--- program BumperF_C (robot ABB IRB 1300-10/1.15) ---
  Smooth(1)
  Set speed (1000.0 mm/s)
  Set Ref.: BumperF
  Set Tool: Generic Paint Sprayer
  Show Generic Paint Sprayer
  MoveJ 1 to (1571.24, -957.53, 569.46) mm, rotated rx 115.95 ry -6.64 rz -166.63 deg; joints [132.246, 136.209, -181.396, 156.344, 105.383, -115.772, 4593.947, 921.715, 1041.563]
  MoveL 2 to (1571.24, -957.53, 569.46) mm, rotated rx 115.95 ry -6.64 rz -166.63 deg; joints [132.246, 136.209, -181.396, 156.344, 105.383, -115.772, 4593.947, 921.715, 1041.563]
  MoveL 3 to (1545.53, -871.22, 525.99) mm, rotated rx 115.95 ry -6.64 rz -166.63 deg; joints [132.246, 136.209, -181.396, 156.344, 105.383, -115.772, 4568.236, 1008.026, 1085.031]
  MoveL 4 to (1545.53, -871.22, 525.99) mm, rotated rx 115.95 ry -6.64 rz -166.63 deg; joints [132.246, 136.209, -181.396, 156.344, 105.383, -115.772, 4568.236, 1008.026, 1085.031]
  Set speed (200.0 mm/s)
  MoveL 5 to (1567.25, -870.44, 513.69) mm, rotated rx 114.53 ry -6.57 rz -165.92 deg; joints [131.765, 135.013, -181.396, 155.74, 105.383, -114.904, 4591.602, 1008.066, 1094.602]
  MoveL 6 to (1592.89, -869.13, 497.74) mm, rotated rx 110.93 ry -5.65 rz -165.57 deg; joints [130.698, 131.085, -181.396, 155.714, 105.383, -112.016, 4607.617, 1008.267, 1096.076]
  MoveL 7 to (1616.69, -868.87, 477.59) mm, rotated rx 107.37 ry -5.12 rz -164.07 deg; joints [129.332, 127.093, -181.396, 154.983, 104.902, -109.292, 4628.08, 1008.268, 1100]
  MoveL 8 to (1638.67, -867.82, 457.97) mm, rotated rx 105.23 ry -4.69 rz -163.28 deg; joints [128.5, 123.788, -181.396, 154.835, 103.912, -107.249, 4645.228, 1008.269, 1099.981]
  MoveL 9 to (1659.86, -866.51, 437.3) mm, rotated rx 104.04 ry -4.24 rz -163.53 deg; joints [128.5, 121.033, -181.396, 155.103, 102.7, -105.772, 4660.763, 1003.997, 1100]
  MoveL 10 to (1680.53, -864.68, 416.9) mm, rotated rx 102.62 ry -4.06 rz -162.44 deg; joints [127.494, 118.2, -181.396, 154.969, 101.395, -104.09, 4676.396, 1006.029, 1100]
  MoveL 11 to (1700.41, -862.07, 396.49) mm, rotated rx 100.96 ry -3.66 rz -161.77 deg; joints [126.76, 115.027, -181.132, 154.969, 100.379, -102.383, 4689.707, 1006.022, 1100]
  MoveL 12 to (1721.6, -858.14, 377.92) mm, rotated rx 98.48 ry -2.82 rz -161.72 deg; joints [126.547, 111.062, -179.997, 154.969, 100.379, -100.648, 4704.908, 1003.768, 1100]
  MoveL 13 to (1729.97, -859.97, 342.08) mm, rotated rx 96.18 ry -2.12 rz -161.17 deg; joints [125.885, 105.454, -176.974, 154.97, 100.379, -99.014, 4709.436, 1003.105, 1100]
  MoveL 14 to (1729.45, -862.07, 324.55) mm, rotated rx 95.53 ry -1.83 rz -161.71 deg; joints [126.39, 103.099, -175.393, 154.981, 100.379, -98.605, 4709.436, 996.85, 1100]
  MoveL 15 to (1734.68, -862.07, 305.71) mm, rotated rx 94.94 ry -1.6 rz -162.14 deg; joints [126.39, 100.689, -173.732, 155.4, 100.379, -98.09, 4710.155, 996.383, 1100]
  MoveL 16 to (1743.31, -860.76, 287.4) mm, rotated rx 94.35 ry -1.49 rz -161.17 deg; joints [125.481, 98.526, -173.288, 155.4, 99.369, -97.19, 4712.272, 996.382, 1100]
  MoveL 17 to (1754.56, -857.88, 271.44) mm, rotated rx 93.88 ry -1.28 rz -161.73 deg; joints [125.481, 96.542, -172.176, 155.976, 99.142, -96.642, 4715.904, 996.382, 1100]
  MoveL 18 to (1759.01, -858.14, 245.02) mm, rotated rx 92.82 ry -0.95 rz -161.34 deg; joints [125.066, 92.989, -169.805, 155.975, 99.142, -95.921, 4715.904, 993.682, 1100]
  MoveL 19 to (1756.13, -859.71, 226.97) mm, rotated rx 92.24 ry -0.73 rz -162.03 deg; joints [125.745, 90.661, -168.159, 155.976, 99.142, -95.55, 4711.513, 983.719, 1100]
  MoveL 20 to (1756.92, -860.24, 208.39) mm, rotated rx 91.53 ry -0.48 rz -162.48 deg; joints [126.192, 88.179, -166.477, 155.976, 99.142, -95.085, 4709.215, 974.937, 1100]
  MoveL 21 to (1757.7, -860.24, 190.6) mm, rotated rx 91.06 ry -0.32 rz -163.42 deg; joints [127.122, 85.976, -164.811, 155.976, 99.142, -94.779, 4708.177, 964.459, 1100]
  MoveL 22 to (1758.49, -860.24, 174.38) mm, rotated rx 90.59 ry -0.18 rz -163.41 deg; joints [127.122, 83.931, -163.287, 155.969, 99.142, -94.457, 4705.559, 959.867, 1100]
  MoveL 23 to (1758.75, -860.24, 159.73) mm, rotated rx 90.12 ry -0.03 rz -163.88 deg; joints [127.59, 82.032, -161.91, 155.969, 99.142, -94.134, 4702.574, 951.798, 1100]
  MoveL 24 to (1759.27, -859.97, 146.91) mm, rotated rx 90 ry 0 rz -165.53 deg; joints [129.218, 80.632, -160.641, 155.988, 99.142, -94.048, 4702.574, 938.888, 1100]
  MoveL 25 to (1760.58, -859.71, 136.45) mm, rotated rx 90.12 ry -0.04 rz -162.94 deg; joints [127.222, 79.74, -160.641, 155.454, 98.168, -93.794, 4702.575, 945.045, 1099.999]
  MoveL 26 to (1763.2, -858.93, 129.12) mm, rotated rx 90.71 ry -0.2 rz -164.47 deg; joints [128.117, 79.543, -159.846, 156.101, 98.168, -94.096, 4702.574, 944.116, 1100]
  Set speed (1000.0 mm/s)
  MoveL 27 to (1763.2, -858.93, 129.12) mm, rotated rx 90.71 ry -0.2 rz -164.47 deg; joints [128.117, 79.543, -159.846, 156.101, 98.168, -94.096, 4702.574, 944.116, 1100]
  MoveL 28 to (1789.97, -955.27, 130.36) mm, rotated rx 90.71 ry -0.2 rz -164.47 deg; joints [128.117, 79.543, -159.846, 156.101, 98.168, -94.096, 4729.346, 847.775, 1098.767]
  Set speed (1000.0 mm/s)
  MoveL 29 to (1779.18, -953.4, 138.35) mm, rotated rx 98.16 ry 0.3 rz 177.94 deg; joints [138.476, 85.541, -159.846, 163.825, 98.168, -98.714, 4697.875, 847.774, 1094.184]
  MoveL 30 to (1782.82, -854.48, 124.15) mm, rotated rx 98.16 ry 0.3 rz 177.94 deg; joints [138.575, 84.798, -159.846, 163.754, 97.448, -98.53, 4697.874, 941.635, 1100]
  MoveL 31 to (1782.82, -854.48, 124.15) mm, rotated rx 98.16 ry 0.3 rz 177.94 deg; joints [138.575, 84.798, -159.846, 163.754, 97.448, -98.53, 4697.874, 941.635, 1100]
  Set speed (200.0 mm/s)
  MoveL 32 to (1786.22, -852.91, 135.66) mm, rotated rx 96.28 ry 0.04 rz 179.68 deg; joints [137.268, 84.574, -160.749, 163.124, 97.823, -97.175, 4697.874, 941.635, 1100]
  MoveL 33 to (1790.67, -851.08, 147.7) mm, rotated rx 98.11 ry -0.22 rz -178.44 deg; joints [135.583, 84.574, -160.749, 163.124, 96.101, -97.893, 4702.805, 954.913, 1071.274]
  MoveL 34 to (1796.68, -848.72, 159.47) mm, rotated rx 98.74 ry -0.53 rz -176.58 deg; joints [133.77, 84.574, -160.749, 163.124, 95.404, -97.953, 4707.715, 968.876, 1052.965]
  MoveL 35 to (1802.7, -846.37, 171.77) mm, rotated rx 98.62 ry -0.68 rz -175.51 deg; joints [133.516, 84.592, -160.749, 162.287, 95.39, -97.953, 4720.878, 970.014, 1041.305]
  MoveL 36 to (1809.24, -843.75, 184.32) mm, rotated rx 99.8 ry -0.99 rz -174.27 deg; joints [132.393, 84.592, -160.749, 162.287, 94.205, -98.297, 4727.536, 980.866, 1017.452]
  MoveL 37 to (1816.57, -840.61, 197.4) mm, rotated rx 100.78 ry -1.11 rz -174.17 deg; joints [132.393, 84.592, -160.749, 162.298, 93.3, -98.698, 4735.96, 985.217, 995.643]
  MoveL 38 to (1824.41, -837.21, 211.01) mm, rotated rx 101.64 ry -1.18 rz -174.28 deg; joints [132.393, 84.592, -160.749, 162.521, 92.536, -99.039, 4742.893, 990.437, 974.508]
  MoveL 39 to (1824.41, -837.21, 211.01) mm, rotated rx 93.53 ry -1.19 rz -161.37 deg; joints [123.735, 79.476, -160.749, 157.598, 94.418, -94.055, 4742.893, 990.436, 988.777]
  MoveL 40 to (1820.23, -837.21, 231.94) mm, rotated rx 93.35 ry -1.2 rz -160.31 deg; joints [123.243, 79.476, -160.872, 157.02, 94.418, -93.99, 4742.894, 992.111, 969.266]
  MoveL 41 to (1820.23, -837.21, 231.94) mm, rotated rx 101.71 ry -1.43 rz -173.11 deg; joints [131.794, 84.617, -160.872, 161.941, 92.215, -98.959, 4742.894, 992.113, 952.179]
  MoveL 42 to (1829.38, -833.03, 246.59) mm, rotated rx 102.88 ry -1.89 rz -171.78 deg; joints [130.559, 84.617, -160.872, 161.941, 90.966, -99.177, 4752.022, 1006.027, 925.876]
  MoveL 43 to (1839.06, -828.32, 260.98) mm, rotated rx 103.06 ry -1.91 rz -171.82 deg; joints [130.559, 84.617, -160.872, 162.004, 90.806, -99.242, 4761.37, 1011.202, 909.915]
  MoveL 44 to (1849.01, -823.35, 275.1) mm, rotated rx 104.57 ry -2.33 rz -171.12 deg; joints [130.013, 84.617, -160.872, 162.004, 89.294, -99.68, 4772.697, 1022.45, 881.62]
  MoveL 45 to (1863.66, -815.76, 294.46) mm, rotated rx 107.07 ry -3 rz -170.32 deg; joints [129.479, 84.698, -160.872, 162.004, 86.864, -100.462, 4790.854, 1039.487, 839.866]
  MoveL 46 to (1882.49, -804.77, 317.22) mm, rotated rx 109.65 ry -4.19 rz -168.43 deg; joints [127.743, 84.698, -160.872, 162.004, 84.028, -100.823, 4811.061, 1068.912, 791.558]
  MoveL 47 to (1895.83, -796.14, 330.83) mm, rotated rx 113.34 ry -6.41 rz -165.49 deg; joints [124.807, 84.698, -160.872, 162.004, 79.723, -100.879, 4824.82, 1109.926, 740.477]
  MoveL 48 to (1904.47, -789.86, 337.89) mm, rotated rx 116.65 ry -8.76 rz -163.11 deg; joints [122.23, 85.616, -160.872, 162.003, 76.566, -100.879, 4837.457, 1154.33, 710.031]
  MoveL 49 to (1913.1, -783.32, 343.38) mm, rotated rx 120.5 ry -11.96 rz -160.62 deg; joints [119.262, 88.097, -160.872, 162.003, 74.023, -100.879, 4855.125, 1218.718, 694.119]
  MoveL 50 to (1922, -776, 347.57) mm, rotated rx 123.01 ry -13.87 rz -159.75 deg; joints [118.011, 89.326, -160.872, 162.003, 72.107, -100.879, 4869.128, 1258.002, 680.927]
  MoveL 51 to (1931.15, -768.41, 350.45) mm, rotated rx 127.02 ry -16.88 rz -158.94 deg; joints [116.434, 91.393, -160.872, 162.003, 69.207, -100.88, 4887.234, 1316.61, 667.809]
  MoveL 52 to (1940.57, -759.78, 352.02) mm, rotated rx 133.81 ry -20.92 rz -159.59 deg; joints [115.619, 92.398, -160.872, 162.003, 62.545, -100.88, 4909.28, 1386.174, 628.482]
  MoveL 53 to (1949.99, -750.62, 352.54) mm, rotated rx 133.85 ry -22.45 rz -158.32 deg; joints [113.518, 92.645, -160.872, 161.597, 62.116, -99.201, 4909.281, 1414.858, 628.482]
  MoveL 54 to (1959.93, -740.68, 352.54) mm, rotated rx 138.13 ry -26.48 rz -158.22 deg; joints [110.548, 94.884, -160.872, 161.597, 59.126, -97.312, 4911.466, 1494.181, 628.482]
  MoveL 55 to (1970.13, -729.69, 351.76) mm, rotated rx 138.94 ry -28.75 rz -157.27 deg; joints [108.289, 95.245, -160.871, 160.752, 58.015, -95.019, 4911.466, 1532.276, 628.482]
  MoveL 56 to (1980.07, -718.44, 350.97) mm, rotated rx 138.97 ry -29.76 rz -156.64 deg; joints [106.869, 95.245, -160.871, 160.411, 57.708, -93.633, 4911.467, 1554.428, 628.83]
  MoveL 57 to (1989.75, -706.93, 349.92) mm, rotated rx 136.16 ry -29.58 rz -154.64 deg; joints [105.639, 94.385, -160.871, 159.72, 59.288, -92.34, 4911.466, 1550.094, 633.425]
  MoveL 58 to (1998.91, -695.68, 349.4) mm, rotated rx 133.19 ry -28.72 rz -152.89 deg; joints [104.809, 93.375, -160.871, 159.442, 61.115, -91.65, 4911.467, 1539.501, 637.871]
  MoveL 59 to (2007.02, -685.48, 349.66) mm, rotated rx 130.86 ry -27.24 rz -152.11 deg; joints [104.689, 92.218, -160.872, 159.777, 62.539, -91.731, 4911.472, 1524.592, 637.872]
  MoveL 60 to (2014.35, -675.8, 350.97) mm, rotated rx 122.46 ry -23.36 rz -148.07 deg; joints [103.96, 90.632, -160.872, 159.151, 69.542, -91.731, 4911.472, 1473.431, 675.241]
  MoveL 61 to (2038.15, -649.11, 345.74) mm, rotated rx 114.17 ry -24.24 rz -137.55 deg; joints [97.018, 85.715, -160.872, 155.117, 71.4, -85.824, 4911.471, 1473.426, 679.245]
  MoveL 62 to (2051.49, -633.42, 343.12) mm, rotated rx 112.8 ry -23.19 rz -136.86 deg; joints [96.789, 84.623, -160.872, 155.117, 71.99, -85.767, 4922.042, 1473.425, 681.907]
  MoveL 63 to (2063.79, -619.03, 341.03) mm, rotated rx 110.74 ry -21.37 rz -136.1 deg; joints [96.739, 82.665, -160.872, 155.117, 72.722, -85.767, 4931.522, 1459.566, 682.288]
  MoveL 64 to (2075.04, -605.69, 338.68) mm, rotated rx 110.8 ry -22.47 rz -134.83 deg; joints [94.985, 82.747, -160.872, 155.117, 72.306, -84.714, 4932.35, 1484.471, 682.288]
  MoveL 65 to (2085.24, -593.13, 336.58) mm, rotated rx 111.8 ry -23.63 rz -134.94 deg; joints [94.569, 83.495, -160.872, 155.119, 71.667, -84.319, 4940.301, 1511.538, 682.287]
  MoveL 66 to (2094.4, -581.62, 334.49) mm, rotated rx 111.31 ry -24.25 rz -133.53 deg; joints [92.994, 83.3, -160.872, 155.016, 71.667, -83.386, 4940.301, 1528.356, 684.409]
  MoveL 67 to (2102.51, -570.63, 332.4) mm, rotated rx 109.4 ry -23.08 rz -131.93 deg; joints [92.04, 82.56, -160.874, 155.016, 73.082, -83.386, 4943.467, 1528.189, 695.451]
  MoveL 68 to (2110.1, -560.43, 330.04) mm, rotated rx 108.78 ry -24.16 rz -129.72 deg; joints [90.063, 82.505, -160.874, 154.429, 73.082, -82.108, 4943.467, 1549.13, 699.124]
  MoveL 69 to (2116.64, -550.75, 327.16) mm, rotated rx 108.04 ry -24.56 rz -128.09 deg; joints [88.633, 82.011, -160.874, 154.121, 73.082, -81.209, 4943.468, 1560.135, 701.179]
  MoveL 70 to (2122.13, -542.64, 323.24) mm, rotated rx 107.35 ry -27.97 rz -123.66 deg; joints [85.357, 82.011, -160.874, 151.788, 72.164, -77.874, 4943.468, 1597.347, 702.069]
  MoveL 71 to (2126.32, -536.1, 317.48) mm, rotated rx 104.82 ry -29.37 rz -118.34 deg; joints [82.164, 80.426, -160.874, 149.535, 72.164, -74.977, 4943.468, 1609.549, 706.168]
  MoveL 72 to (2128.93, -531.65, 312.25) mm, rotated rx 101.45 ry -27.26 rz -113.85 deg; joints [79.937, 78.849, -160.874, 148.686, 74.318, -74.977, 4943.468, 1602.173, 725.352]
  MoveL 73 to (2128.93, -531.65, 312.25) mm, rotated rx 126.84 ry -33.58 rz -143.56 deg; joints [92.503, 91.12, -160.874, 157.962, 63.217, -81.642, 4943.468, 1719.806, 680.931]
  MoveL 74 to (2132.86, -524.59, 312.51) mm, rotated rx 131.8 ry -39.39 rz -144.63 deg; joints [90.442, 93.308, -160.873, 155.312, 59.914, -77.41, 4943.469, 1794.525, 680.931]
  MoveL 75 to (2138.61, -511.5, 310.94) mm, rotated rx 142.1 ry -48.23 rz -149.86 deg; joints [88.012, 93.628, -151.887, 151.963, 59.913, -73.067, 4943.469, 1959.558, 680.933]
  MoveL 76 to (2145.41, -491.62, 307.54) mm, rotated rx 148.42 ry -53.14 rz -153.81 deg; joints [86.275, 93.628, -151.373, 148.126, 56.76, -67.236, 4943.47, 2030.159, 680.933]
  MoveL 77 to (2152.48, -464.94, 303.62) mm, rotated rx 151.46 ry -56.88 rz -155.51 deg; joints [84.483, 93.628, -151.372, 144.702, 55.943, -62.304, 4943.47, 2082.544, 691.657]
  MoveL 78 to (2159.28, -432.5, 300.48) mm, rotated rx 157.96 ry -60.16 rz -160.65 deg; joints [83.237, 93.628, -150.316, 141.632, 54.856, -57.784, 4943.47, 2154.516, 700.89]
  MoveL 79 to (2166.08, -389.07, 298.39) mm, rotated rx 162.71 ry -60.68 rz -164.82 deg; joints [83.006, 93.628, -148.348, 141.49, 54.655, -57.243, 4943.475, 2227.842, 705.926]
  MoveL 80 to (2172.36, -330.47, 297.08) mm, rotated rx 166.98 ry -61.73 rz -168.49 deg; joints [82.432, 93.628, -147.038, 140.505, 54.605, -55.672, 4943.475, 2310.718, 713.199]
  MoveL 81 to (2178.12, -262.97, 296.29) mm, rotated rx 166.1 ry -61.33 rz -167.75 deg; joints [82.2, 93.628, -147.375, 141.056, 54.605, -55.884, 4943.475, 2371.713, 711.376]
  MoveL 82 to (2182.83, -193.12, 295.77) mm, rotated rx 169.21 ry -61.46 rz -170.5 deg; joints [82.021, 93.628, -146.721, 140.72, 54.052, -55.086, 4943.475, 2456.324, 712.371]
  MoveL 83 to (2185.96, -124.84, 295.51) mm, rotated rx 172.94 ry -62.25 rz -173.75 deg; joints [81.639, 93.628, -145.665, 139.712, 54.052, -53.733, 4943.475, 2544.405, 718.894]
  MoveL 84 to (2187.8, -61.27, 295.51) mm, rotated rx 174.69 ry -62.34 rz -175.3 deg; joints [81.557, 93.628, -144.992, 139.539, 54.052, -53.476, 4943.475, 2618.074, 721.416]
  MoveL 85 to (2189.1, -0.05, 295.51) mm, rotated rx -177.26 ry -62.45 rz 177.57 deg; joints [81.557, 93.628, -143.265, 137.966, 52.878, -51.455, 4943.475, 2717.714, 728.542]
  MoveL 86 to (2187.8, 61.17, 295.51) mm, rotated rx -173.75 ry -62.29 rz 174.47 deg; joints [81.71, 93.628, -142.223, 137.399, 52.478, -50.92, 4943.474, 2797.79, 733.234]
  MoveL 87 to (2185.96, 124.74, 295.51) mm, rotated rx -170.29 ry -62.04 rz 171.41 deg; joints [81.906, 93.628, -140.949, 136.945, 52.22, -50.617, 4943.472, 2881.625, 739.388]
  MoveL 88 to (2182.83, 193.28, 295.77) mm, rotated rx -166.22 ry -61.1 rz 167.88 deg; joints [82.416, 93.628, -139.453, 136.732, 51.343, -50.616, 4943.472, 2975.922, 744.195]
  MoveL 89 to (2178.12, 262.87, 296.29) mm, rotated rx -163.59 ry -60.95 rz 165.56 deg; joints [82.676, 93.628, -138.26, 136.285, 51.343, -50.526, 4943.472, 3062.322, 751.37]
  MoveL 90 to (2172.36, 330.37, 297.08) mm, rotated rx -163.15 ry -61.13 rz 165.14 deg; joints [82.913, 93.628, -138.152, 135.936, 51.343, -50.479, 4943.471, 3131.981, 752.579]
  MoveL 91 to (2166.08, 388.97, 298.39) mm, rotated rx -155.06 ry -58.82 rz 158.3 deg; joints [83.805, 93.628, -134.575, 135.497, 49.863, -50.479, 4943.471, 3246.959, 770.044]
  MoveL 92 to (2159.28, 432.4, 300.48) mm, rotated rx -150.95 ry -57.83 rz 154.82 deg; joints [84.274, 93.628, -132.455, 135.037, 49.517, -50.479, 4943.457, 3320.012, 783.091]
  MoveL 93 to (2152.48, 465.1, 303.62) mm, rotated rx -144.6 ry -53.45 rz 150.28 deg; joints [85.716, 93.628, -130.007, 135.037, 45.48, -50.342, 4943.456, 3409.512, 793.219]
  MoveL 94 to (2145.41, 491.52, 307.54) mm, rotated rx -142.77 ry -49.52 rz 149.98 deg; joints [86.332, 93.736, -130.007, 136.122, 41.249, -50.342, 4923.205, 3464.712, 785.161]
  MoveL 95 to (2138.61, 511.67, 310.94) mm, rotated rx -140.46 ry -46.77 rz 148.98 deg; joints [87.496, 93.756, -129.75, 136.122, 37.777, -50.276, 4923.205, 3511.087, 785.16]
  MoveL 96 to (2132.86, 524.49, 312.51) mm, rotated rx -133.08 ry -41.17 rz 144.86 deg; joints [88.774, 93.756, -125.065, 136.122, 33.797, -50.263, 4923.205, 3605.485, 833.592]
  MoveL 97 to (2128.93, 531.55, 312.25) mm, rotated rx -126.84 ry -33.58 rz 143.56 deg; joints [90.862, 93.756, -122.789, 136.122, 25.461, -49.709, 4923.205, 3689.917, 878.711]
  MoveL 98 to (2128.93, 531.55, 312.25) mm, rotated rx -100.25 ry -7.61 rz 109.92 deg; joints [121.937, 78.369, -126.316, 15.017, 36.087, 78.198, 5588.694, 3468.859, 878.521]
  MoveL 99 to (2126.32, 536, 317.48) mm, rotated rx -104.1 ry -29.19 rz 117.26 deg; joints [117.367, 96.341, -169.247, 16.72, 48.145, 64.164, 5423.205, 3346.609, 878.683]
  MoveL 100 to (2122.13, 542.54, 323.24) mm, rotated rx -105.97 ry -28.47 rz 120.97 deg; joints [117.367, 96.341, -169.247, 12.679, 46.638, 66.806, 5394.89, 3369.672, 861.092]
  MoveL 101 to (2116.64, 550.65, 327.16) mm, rotated rx -107.55 ry -25.57 rz 126.23 deg; joints [117.365, 96.872, -169.247, 5.15, 45.601, 72.802, 5349.984, 3412.333, 858.641]
  MoveL 102 to (2110.1, 560.33, 330.04) mm, rotated rx -108.36 ry -23.05 rz 130.28 deg; joints [117.365, 97.148, -169.622, -1.121, 45.94, 77.838, 5308.188, 3445.265, 858.641]
  MoveL 103 to (2102.51, 570.53, 332.4) mm, rotated rx -108.16 ry -21.99 rz 131.22 deg; joints [117.365, 97.148, -169.622, -2.931, 46.544, 79.449, 5290.898, 3463.725, 860.533]
  MoveL 104 to (2094.4, 581.52, 334.49) mm, rotated rx -112.03 ry -24.25 rz 134.57 deg; joints [117.365, 97.148, -169.622, -4.906, 42.427, 79.382, 5264.861, 3465.093, 824.183]
  MoveL 105 to (2085.24, 593.29, 336.58) mm, rotated rx -112.13 ry -23.27 rz 135.83 deg; joints [117.365, 97.206, -169.702, -7.138, 42.788, 81.232, 5243.276, 3484.334, 824.183]
  MoveL 106 to (2075.04, 605.59, 338.68) mm, rotated rx -109.09 ry -20.54 rz 134.6 deg; joints [117.942, 97.207, -169.702, -8.433, 46.502, 83.15, 5241.183, 3509.289, 851.703]
  MoveL 107 to (2063.79, 618.93, 341.03) mm, rotated rx -110.74 ry -21.37 rz 136.11 deg; joints [117.941, 97.207, -169.702, -9.617, 44.796, 83.448, 5220.921, 3519.123, 834.664]
  MoveL 108 to (2051.49, 633.32, 343.12) mm, rotated rx -112.8 ry -23.16 rz 136.91 deg; joints [118.362, 97.207, -169.702, -9.734, 42.342, 82.526, 5213.697, 3519.123, 812.954]
  MoveL 109 to (2038.15, 649.01, 345.74) mm, rotated rx -114.2 ry -23.4 rz 138.54 deg; joints [118.362, 97.207, -169.702, -11.45, 41.13, 83.478, 5189.149, 3533.479, 799.64]
  MoveL 110 to (2014.35, 675.7, 350.97) mm, rotated rx -123.67 ry -27.39 rz 145.37 deg; joints [118.362, 100.052, -169.702, -17.048, 29.191, 86.118, 5142.169, 3533.473, 756.191]
  MoveL 111 to (2007.02, 685.38, 349.66) mm, rotated rx -129.78 ry -26.88 rz 151.5 deg; joints [118.361, 102.105, -169.702, -29.591, 23.106, 96.935, 5097.394, 3533.473, 745.089]
  MoveL 112 to (1998.91, 695.84, 349.4) mm, rotated rx -134.96 ry -27.94 rz 154.87 deg; joints [118.362, 104.566, -169.702, -40.535, 16.934, 107.101, 5081.009, 3524.437, 745.027]
  MoveL 113 to (1989.75, 706.83, 349.92) mm, rotated rx -135.77 ry -28.84 rz 154.84 deg; joints [118.599, 104.566, -169.702, -39.809, 15.836, 106.09, 5081.008, 3525.47, 739.705]
  MoveL 114 to (1980.07, 718.34, 350.97) mm, rotated rx -137.63 ry -29.46 rz 155.84 deg; joints [118.599, 104.853, -169.702, -43.067, 14.024, 109.061, 5070.617, 3525.467, 732.328]
  MoveL 115 to (1970.13, 729.59, 351.76) mm, rotated rx -137.6 ry -27.86 rz 156.89 deg; joints [118.702, 104.851, -169.702, -48.91, 15.339, 114.706, 5045.317, 3542.967, 732.328]
  MoveL 116 to (1959.93, 740.58, 352.54) mm, rotated rx -137.33 ry -25.27 rz 158.52 deg; joints [118.819, 104.799, -169.702, -55.944, 17.838, 121.432, 5009.494, 3564.603, 734.131]
  MoveL 117 to (1949.99, 750.78, 352.54) mm, rotated rx -135.75 ry -22.51 rz 159.55 deg; joints [118.87, 104.794, -169.702, -58.879, 21.266, 124.214, 4975.283, 3593.366, 745.656]
  MoveL 118 to (1940.57, 759.94, 352.02) mm, rotated rx -132.32 ry -19.53 rz 159.84 deg; joints [118.87, 104.805, -169.702, -57.999, 25.87, 123.334, 4944.52, 3631.825, 770.684]
  MoveL 119 to (1931.15, 768.31, 350.45) mm, rotated rx -125.59 ry -15.57 rz 159.44 deg; joints [118.872, 104.805, -169.702, -54.022, 33.33, 119.439, 4914.242, 3687.634, 823.647]
  MoveL 120 to (1922, 776.16, 347.57) mm, rotated rx -122.37 ry -12.62 rz 160.98 deg; joints [120.106, 105.786, -171.045, -56.102, 38.789, 119.815, 4891.208, 3703.918, 865.204]
  MoveL 121 to (1913.1, 783.22, 343.38) mm, rotated rx -118.52 ry -10.68 rz 161.17 deg; joints [122.15, 107.812, -173.857, -56.247, 44.118, 117.831, 4891.207, 3706.572, 920.695]
  MoveL 122 to (1904.47, 789.76, 337.89) mm, rotated rx -114.98 ry -8.12 rz 163.14 deg; joints [125.003, 107.808, -173.858, -60.282, 50.047, 118.539, 4889.848, 3706.573, 961.367]
  MoveL 123 to (1895.83, 796.04, 330.83) mm, rotated rx -111.51 ry -5.54 rz 166.23 deg; joints [126.979, 107.837, -173.899, -64.217, 56.027, 119.193, 4868.359, 3706.573, 1004.927]
  MoveL 124 to (1882.49, 804.68, 317.22) mm, rotated rx -109.07 ry -4.29 rz 167.78 deg; joints [128.581, 107.838, -173.899, -66.332, 59.756, 119.034, 4855.913, 3706.573, 1042.723]
  MoveL 125 to (1863.66, 815.66, 294.46) mm, rotated rx -105.98 ry -2.95 rz 169.8 deg; joints [130.272, 107.838, -173.899, -68.62, 64.249, 118.586, 4834.611, 3706.573, 1095.868]
  MoveL 126 to (1849.01, 823.51, 275.1) mm, rotated rx -104.09 ry -2.33 rz 170.81 deg; joints [130.355, 105.02, -173.899, -67.719, 67.486, 115.138, 4802.741, 3706.574, 1100]
  MoveL 127 to (1839.06, 828.22, 260.98) mm, rotated rx -103.1 ry -1.96 rz 171.62 deg; joints [130.355, 102.973, -173.899, -67.412, 69.506, 112.896, 4778.483, 3703.896, 1100]
  MoveL 128 to (1829.38, 832.93, 246.59) mm, rotated rx -102.72 ry -1.85 rz 171.86 deg; joints [130.355, 101.399, -173.899, -66.996, 70.557, 111.244, 4761.166, 3702.57, 1100]
  MoveL 129 to (1820.23, 837.38, 231.94) mm, rotated rx -101.39 ry -1.37 rz 173.22 deg; joints [130.355, 98.949, -173.899, -67.213, 73.194, 108.642, 4730.295, 3695.409, 1100]
  MoveL 130 to (1811.6, 841.3, 217.55) mm, rotated rx -100.83 ry -1.21 rz 173.68 deg; joints [130.355, 97.17, -173.898, -67.051, 74.53, 106.798, 4710.472, 3690.876, 1100]
  MoveL 131 to (1804.27, 844.44, 203.42) mm, rotated rx -99.58 ry -0.85 rz 174.97 deg; joints [130.355, 94.672, -172.725, -67.719, 76.533, 105.253, 4686.599, 3686.562, 1099.999]
  MoveL 132 to (1797.73, 847.32, 189.56) mm, rotated rx -98.67 ry -0.72 rz 175.26 deg; joints [130.355, 92.527, -171.328, -67.654, 77.698, 104.177, 4674.566, 3686.562, 1100]
  MoveL 133 to (1791.71, 849.67, 176.21) mm, rotated rx -97.52 ry -0.56 rz 175.77 deg; joints [130.355, 90.189, -169.438, -67.837, 79.01, 103.309, 4662.082, 3686.561, 1100]
  MoveL 134 to (1786.22, 851.77, 163.39) mm, rotated rx -96.75 ry -0.35 rz 177.02 deg; joints [130.355, 88.16, -167.134, -68.975, 79.879, 103.424, 4646.519, 3686.561, 1100]
  MoveL 135 to (1780.99, 853.6, 150.57) mm, rotated rx -96.72 ry -0.25 rz 177.84 deg; joints [130.355, 86.792, -165.498, -69.827, 80.013, 103.801, 4634.934, 3686.561, 1100]
  MoveL 136 to (1776.02, 855.43, 138.28) mm, rotated rx -97.31 ry -0.15 rz 178.83 deg; joints [130.199, 86.008, -164.453, -70.824, 79.637, 104.515, 4620.637, 3686.561, 1100]
  Set speed (1000.0 mm/s)
  MoveL 137 to (1776.02, 855.43, 138.28) mm, rotated rx -97.31 ry -0.15 rz 178.83 deg; joints [130.199, 86.008, -164.453, -70.824, 79.637, 104.515, 4620.637, 3686.561, 1100]
  MoveL 138 to (1778.07, 954.59, 151.01) mm, rotated rx -97.31 ry -0.15 rz 178.83 deg; joints [130.199, 86.008, -164.453, -70.824, 79.637, 104.515, 4622.694, 3785.727, 1087.273]
  Set speed (1000.0 mm/s)
  MoveL 139 to (1808.49, 946.12, 127.52) mm, rotated rx -90.28 ry -0.17 rz 148.43 deg; joints [129.033, 79.118, -164.453, -37.565, 85.971, 92.833, 4884.487, 3785.726, 1100]
  MoveL 140 to (1756.13, 860.92, 127.03) mm, rotated rx -90.28 ry -0.17 rz 148.43 deg; joints [129.033, 79.068, -164.387, -37.566, 85.959, 92.843, 4832.141, 3700.553, 1100]
  MoveL 141 to (1756.13, 860.92, 127.03) mm, rotated rx -90.28 ry -0.17 rz 148.43 deg; joints [129.033, 79.068, -164.387, -37.566, 85.959, 92.843, 4832.141, 3700.553, 1100]
  Set speed (200.0 mm/s)
  MoveL 142 to (1755.35, 861.18, 142.2) mm, rotated rx -89.73 ry 0.15 rz 149.83 deg; joints [129.033, 79.823, -164.388, -38.967, 86.078, 93.416, 4822.58, 3707.684, 1098.225]
  MoveL 143 to (1754.3, 861.71, 158.16) mm, rotated rx -91.03 ry -0.62 rz 148.95 deg; joints [129.033, 78.833, -163.076, -38.196, 84.269, 93.535, 4830.145, 3707.674, 1058.331]
  MoveL 144 to (1752.47, 862.23, 174.91) mm, rotated rx -92.22 ry -1.36 rz 148.58 deg; joints [129.033, 77.963, -161.93, -37.903, 82.624, 93.64, 4832.255, 3707.563, 1019.854]
  MoveL 145 to (1750.12, 862.75, 193.22) mm, rotated rx -92.85 ry -1.8 rz 147.69 deg; joints [129.033, 77.382, -161.169, -37.055, 81.659, 93.607, 4838.475, 3706.721, 988.749]
  MoveL 146 to (1746.45, 863.54, 212.84) mm, rotated rx -94.48 ry -2.91 rz 147.03 deg; joints [129.033, 76.121, -159.522, -36.478, 79.343, 93.646, 4841.659, 3705.121, 938.551]
  MoveL 147 to (1741.74, 864.32, 234.03) mm, rotated rx -95.15 ry -3.34 rz 147.13 deg; joints [129.04, 75.664, -158.928, -36.626, 78.443, 93.712, 4836.3, 3705.121, 905.494]
  MoveL 148 to (1735.73, 865.37, 256.79) mm, rotated rx -97.44 ry -4.81 rz 147.32 deg; joints [129.04, 74.055, -156.847, -36.901, 75.36, 93.907, 4829.618, 3702.339, 842.017]
  MoveL 149 to (1728.14, 866.42, 280.86) mm, rotated rx -98.87 ry -5.68 rz 147.6 deg; joints [129.04, 73.076, -155.588, -37.228, 73.484, 94.072, 4820.151, 3700.418, 793.148]
  MoveL 150 to (1718.98, 867.46, 305.97) mm, rotated rx -100.37 ry -6.31 rz 149.01 deg; joints [129.04, 72.307, -154.602, -38.728, 71.812, 94.585, 4798.594, 3699.518, 745.657]
  MoveL 151 to (1708, 868.77, 331.09) mm, rotated rx -101.98 ry -7.27 rz 149.2 deg; joints [129.067, 71.173, -153.156, -38.984, 69.715, 94.797, 4787.11, 3695.693, 692.782]
  MoveL 152 to (1695.18, 870.08, 356.2) mm, rotated rx -104.66 ry -8.53 rz 150.44 deg; joints [129.067, 69.501, -151.034, -40.362, 66.539, 95.52, 4764.249, 3688.816, 625.271]
  MoveL 153 to (1680.79, 871.13, 380.27) mm, rotated rx -107.37 ry -9.65 rz 151.83 deg; joints [129.067, 67.833, -148.932, -41.928, 63.447, 96.434, 4738.607, 3679.945, 559.722]
  MoveL 154 to (1664.57, 872.43, 403.29) mm, rotated rx -110.26 ry -10.66 rz 153.37 deg; joints [129.067, 66.074, -146.727, -43.757, 60.286, 97.612, 4709.613, 3668.958, 494.072]
  MoveL 155 to (1646.78, 873.74, 425.27) mm, rotated rx -111.51 ry -11.45 rz 153.27 deg; joints [129.568, 65.251, -145.7, -44.169, 58.711, 97.776, 4698.886, 3659.227, 452.239]
  MoveL 156 to (1627.68, 875.05, 445.94) mm, rotated rx -116.57 ry -12.63 rz 156.39 deg; joints [129.568, 62.273, -142.003, -48.212, 53.661, 100.655, 4652.997, 3634.303, 362.586]
  MoveL 157 to (1607.01, 876.36, 465.3) mm, rotated rx -121.2 ry -14.2 rz 157.95 deg; joints [129.834, 59.147, -138.156, -50.902, 48.704, 102.937, 4623.002, 3602.462, 278.009]
  MoveL 158 to (1585.04, 877.4, 483.35) mm, rotated rx -123.01 ry -14.13 rz 159.4 deg; joints [129.834, 58.182, -136.974, -53.177, 47.297, 104.716, 4587.225, 3592.257, 239.187]
  MoveL 159 to (1562.02, 878.45, 499.83) mm, rotated rx -126.91 ry -13.64 rz 162.56 deg; joints [129.834, 56.118, -134.454, -58.637, 44.608, 109.178, 4532.723, 3567.214, 180.331]
  MoveL 160 to (1537.16, 879.24, 514.74) mm, rotated rx -129.96 ry -13.55 rz 164.37 deg; joints [129.834, 54.196, -132.118, -62.413, 42.314, 112.594, 4489.195, 3544.02, 130.207]
  MoveL 161 to (1511.79, 880.02, 528.35) mm, rotated rx -131.91 ry -13.23 rz 165.7 deg; joints [129.834, 53.019, -130.692, -65.342, 41.109, 115.235, 4449.329, 3528.97, 95.816]
  MoveL 162 to (1496.35, 880.54, 535.15) mm, rotated rx -132.2 ry -12.2 rz 166.87 deg; joints [129.834, 53.299, -130.692, -67.741, 41.65, 117.21, 4421.818, 3531.052, 92.371]
  Set speed (1000.0 mm/s)
  MoveL 163 to (1496.35, 880.54, 535.15) mm, rotated rx -132.2 ry -12.2 rz 166.87 deg; joints [129.834, 53.299, -130.692, -67.741, 41.65, 117.21, 4421.818, 3531.052, 92.371]
  MoveL 164 to (1527, 949.47, 600.8) mm, rotated rx -132.2 ry -12.2 rz 166.87 deg; joints [129.834, 53.299, -130.692, -67.741, 41.65, 117.21, 4452.47, 3599.975, 26.72]
  Set speed (1000.0 mm/s)
  MoveL 165 to (1587.92, 958.15, 549.01) mm, rotated rx -102.23 ry 17.96 rz 168.04 deg; joints [85.247, 75.154, -172.556, -15.527, 95.973, 109.606, 3959.067, 3839.998, 624.018]
  MoveL 166 to (1574.05, 861.18, 528.87) mm, rotated rx -102.23 ry 17.96 rz 168.04 deg; joints [85.247, 75.154, -172.556, -15.527, 95.973, 109.606, 3945.197, 3743.035, 644.162]
  MoveL 167 to (1574.05, 861.18, 528.87) mm, rotated rx -102.23 ry 17.96 rz 168.04 deg; joints [85.247, 75.154, -172.556, -15.527, 95.973, 109.606, 3945.197, 3743.035, 644.162]
  Set speed (200.0 mm/s)
  MoveL 168 to (1582.94, 860.92, 524.16) mm, rotated rx -99.22 ry 18.11 rz 166.27 deg; joints [85.247, 75.154, -172.556, -12.897, 98.564, 108.56, 3978.942, 3749.725, 673.617]
  MoveL 169 to (1601, 858.31, 517.62) mm, rotated rx -101.62 ry 18.6 rz 170.82 deg; joints [85.247, 75.154, -172.557, -18.164, 96.702, 109.516, 3948.452, 3733.48, 663.003]
  MoveL 170 to (1617.22, 859.88, 502.18) mm, rotated rx -100.08 ry 18.75 rz 170.85 deg; joints [85.247, 75.154, -172.556, -17.754, 98.04, 108.926, 3968.868, 3736.767, 691.409]
  MoveL 171 to (1635.27, 859.61, 488.06) mm, rotated rx -97.66 ry 19.02 rz 170.97 deg; joints [85.247, 75.154, -172.493, -17.2, 100.097, 108.057, 3992.85, 3738.739, 725.96]
  MoveL 172 to (1656.46, 858.31, 471.58) mm, rotated rx -95.1 ry 19.33 rz 171.2 deg; joints [85.247, 75.154, -172.404, -16.733, 102.274, 107.18, 4019.475, 3738.739, 764.218]
  MoveL 173 to (1678.17, 856.21, 453.79) mm, rotated rx -91.71 ry 19.73 rz 170.17 deg; joints [85.247, 75.154, -172.404, -14.777, 105.322, 106.175, 4060.772, 3739.258, 811.005]
  MoveL 174 to (1700.67, 853.6, 435.47) mm, rotated rx -90.06 ry 19.99 rz 170.5 deg; joints [85.247, 75.154, -171.85, -14.635, 106.278, 105.801, 4085.023, 3739.258, 842.776]
  MoveL 175 to (1723.69, 850.2, 417.42) mm, rotated rx -88.96 ry 20.14 rz 171.84 deg; joints [84.269, 75.154, -170.835, -14.635, 106.278, 105.692, 4088.131, 3738.545, 868.777]
  MoveL 176 to (1746.98, 845.75, 400.15) mm, rotated rx -86.74 ry 20.53 rz 170.67 deg; joints [84.269, 75.172, -170.361, -12.791, 107.864, 105.333, 4128.741, 3738.545, 904.83]
  MoveL 177 to (1746.98, 845.75, 400.15) mm, rotated rx -100.04 ry 13.11 rz 143.03 deg; joints [84.269, 75.172, -172.274, 11.306, 95.041, 107.735, 4349.929, 3738.545, 769.692]
  MoveL 178 to (1745.15, 852.55, 362.22) mm, rotated rx -101.97 ry 11.95 rz 143.48 deg; joints [84.269, 74.5, -172.275, 10.388, 93.508, 107.75, 4340.519, 3738.545, 781.412]
  MoveL 179 to (1754.3, 853.07, 330.57) mm, rotated rx -90.02 ry 19.99 rz 146.7 deg; joints [84.269, 74.5, -171.915, 10.873, 107.107, 108.909, 4350.239, 3738.546, 942.781]
  MoveL 180 to (1749.33, 856.21, 316.96) mm, rotated rx -92.02 ry 18.69 rz 145.18 deg; joints [84.269, 74.5, -172.519, 11.689, 105.408, 108.899, 4353.587, 3738.545, 936.348]
  MoveL 181 to (1746.98, 857.78, 305.97) mm, rotated rx -90.99 ry 19.37 rz 145.61 deg; joints [84.269, 74.5, -172.519, 11.65, 106.587, 109.018, 4350.414, 3738.995, 958.271]
  Set speed (1000.0 mm/s)
  MoveL 182 to (1746.98, 857.78, 305.97) mm, rotated rx -90.99 ry 19.37 rz 145.61 deg; joints [84.269, 74.5, -172.519, 11.65, 106.587, 109.018, 4350.414, 3738.995, 958.271]
  MoveL 183 to (1802.98, 940.61, 307.6) mm, rotated rx -90.99 ry 19.37 rz 145.61 deg; joints [84.269, 74.5, -172.519, 11.65, 106.587, 109.018, 4406.42, 3821.825, 956.646]
  Set speed (1000.0 mm/s)
  MoveL 184 to (1854.93, 915.91, 367.18) mm, rotated rx -85.82 ry 20.96 rz 166.98 deg; joints [84.269, 76.29, -170.789, -8.659, 108.209, 105.795, 4272.92, 3821.825, 956.645]
  MoveL 185 to (1829.91, 819.33, 373.99) mm, rotated rx -85.82 ry 20.96 rz 166.98 deg; joints [84.269, 76.29, -170.789, -8.659, 108.209, 105.795, 4247.901, 3725.245, 949.833]
  MoveL 186 to (1829.91, 819.33, 373.99) mm, rotated rx -85.82 ry 20.96 rz 166.98 deg; joints [84.269, 76.29, -170.789, -8.659, 108.209, 105.795, 4247.901, 3725.245, 949.833]
  Set speed (200.0 mm/s)
  MoveL 187 to (1811.6, 824.3, 386.81) mm, rotated rx -87.7 ry 20.42 rz 169.25 deg; joints [84.269, 76.29, -171.258, -11.582, 106.816, 105.823, 4202.812, 3725.245, 920.581]
  MoveL 188 to (1788.57, 830.31, 401.2) mm, rotated rx -87.83 ry 20.39 rz 169.59 deg; joints [84.269, 76.29, -171.387, -11.98, 106.816, 105.784, 4176.319, 3729.768, 905.242]
  MoveL 189 to (1763.46, 836.33, 416.9) mm, rotated rx -89.82 ry 20.03 rz 169.74 deg; joints [84.269, 76.29, -172.379, -12.744, 105.956, 106.078, 4144.305, 3729.768, 873.607]
  MoveL 190 to (1738.6, 841.04, 433.64) mm, rotated rx -91.41 ry 19.75 rz 168.94 deg; joints [84.566, 76.29, -173.41, -12.733, 105.508, 106.333, 4125.714, 3729.768, 844.466]
  MoveL 191 to (1714.54, 844.7, 450.91) mm, rotated rx -93.31 ry 19.44 rz 169.34 deg; joints [84.566, 76.29, -173.856, -13.688, 104.206, 106.732, 4092.481, 3729.768, 811.405]
  MoveL 192 to (1691.25, 847.58, 467.91) mm, rotated rx -94.18 ry 19.22 rz 168.13 deg; joints [85.492, 76.29, -174.698, -13.688, 104.206, 106.748, 4087.977, 3730.076, 787.973]
  MoveL 193 to (1669.28, 850.2, 483.35) mm, rotated rx -97.29 ry 18.85 rz 169.33 deg; joints [85.489, 76.29, -174.698, -15.748, 101.404, 107.626, 4045.754, 3729.073, 745.926]
  MoveL 194 to (1648.87, 852.03, 496.17) mm, rotated rx -97.84 ry 18.61 rz 168.1 deg; joints [86.485, 76.29, -175.289, -15.694, 101.404, 107.536, 4045.754, 3729.983, 728.74]
  MoveL 195 to (1630.56, 853.86, 507.15) mm, rotated rx -99.43 ry 18.6 rz 169.52 deg; joints [86.485, 76.29, -175.289, -17.562, 100.024, 108.024, 4009.856, 3727.192, 704.896]
  MoveL 196 to (1615.65, 854.64, 515.79) mm, rotated rx -100.49 ry 18.29 rz 168.53 deg; joints [87.17, 76.29, -175.659, -17.562, 99.357, 108.178, 4008.221, 3727.192, 687.126]
  MoveL 197 to (1596.81, 855.69, 526.51) mm, rotated rx -100.73 ry 18.45 rz 169.53 deg; joints [87.17, 76.311, -175.659, -18.641, 99.164, 108.269, 3979.53, 3725.629, 675.248]
  MoveL 198 to (1577.97, 856.21, 536.98) mm, rotated rx -101.44 ry 18.09 rz 168.13 deg; joints [87.921, 76.311, -176.166, -18.189, 98.908, 108.231, 3979.53, 3725.629, 658.553]
  Set speed (1000.0 mm/s)
  MoveL 199 to (1577.97, 856.21, 536.98) mm, rotated rx -101.44 ry 18.09 rz 168.13 deg; joints [87.921, 76.311, -176.166, -18.189, 98.908, 108.231, 3979.53, 3725.629, 658.553]
  MoveL 200 to (1592.11, 953.4, 555.83) mm, rotated rx -101.44 ry 18.09 rz 168.13 deg; joints [87.921, 76.311, -176.166, -18.189, 98.908, 108.231, 3993.667, 3822.812, 639.697]
  Set speed (1000.0 mm/s)
  MoveL 201 to (1884.33, 847.56, 483.62) mm, rotated rx -150.84 ry -17.1 rz 170.68 deg; joints [105.146, 51.554, -146.258, -32.636, 33.423, 104.112, 4535.971, 3356.589, 26.72]
  MoveL 202 to (1851.1, 803.63, 400.15) mm, rotated rx -150.84 ry -17.1 rz 170.68 deg; joints [105.146, 51.554, -146.258, -32.637, 33.423, 104.112, 4502.744, 3312.663, 110.186]
  MoveL 203 to (1851.1, 803.63, 400.15) mm, rotated rx -150.84 ry -17.1 rz 170.68 deg; joints [105.146, 51.554, -146.258, -32.637, 33.423, 104.112, 4502.744, 3312.663, 110.186]
  Set speed (200.0 mm/s)
  MoveL 204 to (1871.24, 793.69, 395.97) mm, rotated rx -153.3 ry -26.25 rz 167.46 deg; joints [105.146, 52.249, -146.258, -15.49, 27.628, 89.851, 4615.066, 3278.249, 101.824]
  MoveL 205 to (1889.56, 782.7, 392.31) mm, rotated rx -156.08 ry -27.91 rz 168.27 deg; joints [105.146, 52.249, -146.258, -12.631, 24.891, 87.31, 4644.676, 3242.778, 96.428]
  MoveL 206 to (1906.56, 770.67, 389.17) mm, rotated rx -157.76 ry -26.85 rz 169.54 deg; joints [104.53, 52.548, -146.258, -15.686, 23.326, 90.72, 4643.765, 3225.359, 96.428]
  MoveL 207 to (1922.26, 758.11, 386.55) mm, rotated rx -156.28 ry -24.24 rz 169.77 deg; joints [104.53, 52.548, -146.258, -21.481, 25.253, 95.923, 4635.917, 3228.991, 103.943]
  MoveL 208 to (1937.43, 745.03, 383.93) mm, rotated rx -153.43 ry -24.18 rz 168.42 deg; joints [103.829, 51.726, -146.258, -18.788, 28.546, 93.879, 4646.53, 3228.991, 110.554]
  MoveL 209 to (1952.34, 731.95, 381.58) mm, rotated rx -153.48 ry -24.13 rz 168.47 deg; joints [103.783, 51.69, -146.213, -18.888, 28.512, 94.012, 4660.41, 3215.595, 112.478]
  MoveL 210 to (1966.99, 718.34, 379.49) mm, rotated rx -151.25 ry -24.23 rz 167.31 deg; joints [103.543, 51.666, -146.213, -17.267, 30.465, 92.707, 4678.277, 3218.927, 122.453]
  MoveL 211 to (1981.12, 704.74, 377.39) mm, rotated rx -149.69 ry -25.53 rz 165.86 deg; joints [104.543, 51.669, -146.213, -14.653, 31.481, 89.536, 4718.095, 3211.792, 129.99]
  MoveL 212 to (1994.72, 691.4, 375.3) mm, rotated rx -150.04 ry -26.96 rz 165.36 deg; joints [104.543, 51.625, -146.157, -11.78, 30.853, 87.082, 4745.517, 3192.154, 129.99]
  MoveL 213 to (2014.35, 671.25, 371.9) mm, rotated rx -148.86 ry -27.88 rz 164.22 deg; joints [105.352, 51.627, -146.16, -10.08, 31.703, 84.922, 4784.604, 3175.975, 137.909]
  MoveL 214 to (2033.71, 650.85, 368.76) mm, rotated rx -148.33 ry -28.87 rz 163.42 deg; joints [106.26, 51.649, -146.187, -8.629, 31.995, 82.889, 4823.354, 3154.128, 143.316]
  MoveL 215 to (2046.26, 636.72, 366.67) mm, rotated rx -147.12 ry -29.89 rz 162.14 deg; joints [107.248, 51.649, -146.187, -6.98, 32.886, 80.669, 4858.306, 3142.184, 150.368]
  MoveL 216 to (2059.08, 622.07, 364.84) mm, rotated rx -148.97 ry -31.14 rz 162.72 deg; joints [107.249, 51.649, -146.187, -4.864, 31.173, 78.717, 4878.563, 3111.235, 145.335]
  MoveL 217 to (2071.9, 607.16, 363.01) mm, rotated rx -152.27 ry -31.25 rz 164.75 deg; joints [107.194, 51.649, -146.187, -5.252, 28.346, 78.874, 4883.803, 3073.816, 135.3]
  MoveL 218 to (2084.2, 591.98, 361.17) mm, rotated rx -151 ry -31.15 rz 164 deg; joints [107.183, 52.079, -146.187, -5.299, 29.007, 79.028, 4899.74, 3073.219, 144.364]
  MoveL 219 to (2096.23, 576.55, 359.6) mm, rotated rx -151.95 ry -32.02 rz 164.22 deg; joints [107.183, 52.079, -146.187, -3.494, 28.159, 77.355, 4918.037, 3048.723, 143.14]
  MoveL 220 to (2107.22, 561.64, 358.3) mm, rotated rx -152.65 ry -32.13 rz 164.62 deg; joints [107.184, 52.079, -146.187, -3.323, 27.563, 77.149, 4928.525, 3028.706, 142.159]
  MoveL 221 to (2117.68, 546.46, 356.99) mm, rotated rx -153.56 ry -35.01 rz 164.08 deg; joints [107.184, 51.951, -146.028, 3.404, 26.846, 70.989, 4964.458, 2997.99, 142.159]
  MoveL 222 to (2127.1, 531.55, 355.94) mm, rotated rx -159.57 ry -39.86 rz 166.57 deg; joints [107.184, 51.952, -146.028, 17.145, 23.225, 57.519, 5007.397, 2929.606, 134.914]
  MoveL 223 to (2136, 514.02, 354.9) mm, rotated rx -166.11 ry -42.26 rz 170.55 deg; joints [107.184, 52.015, -146.028, 28.982, 19.978, 45.355, 5029.237, 2865.389, 129.661]
  MoveL 224 to (2144.89, 491.78, 353.59) mm, rotated rx -170.65 ry -43.57 rz 173.52 deg; joints [107.184, 52.124, -146.028, 38.669, 18.335, 35.368, 5046.103, 2813.417, 129.643]
  MoveL 225 to (2153, 464.58, 352.54) mm, rotated rx -172.06 ry -43.46 rz 174.52 deg; joints [106.935, 52.124, -146.028, 41.13, 17.597, 33.025, 5050.111, 2777.966, 129.055]
  MoveL 226 to (2160.33, 431.88, 351.49) mm, rotated rx -178.4 ry -42.89 rz 178.91 deg; joints [106.928, 52.179, -146.028, 54.296, 14.831, 19.315, 5050.112, 2705.18, 125.478]
  MoveL 227 to (2166.87, 388.97, 350.45) mm, rotated rx 179.8 ry -41.02 rz -179.87 deg; joints [106.928, 52.82, -146.028, 59.523, 12.297, 13.832, 5042.081, 2658.61, 125.478]
  MoveL 228 to (2173.41, 330.37, 349.66) mm, rotated rx 179.44 ry -39.92 rz -179.64 deg; joints [106.928, 53.112, -146.028, 60.833, 11.021, 12.448, 5039.768, 2601.216, 125.477]
  MoveL 229 to (2178.9, 262.87, 348.88) mm, rotated rx -177.29 ry -39.65 rz 178.27 deg; joints [106.573, 55.452, -146.028, 58.565, 10.192, 15.083, 5048.702, 2587.392, 142.914]
  MoveL 230 to (2183.35, 193.28, 348.09) mm, rotated rx -178.07 ry -40.16 rz 178.76 deg; joints [106.573, 55.235, -145.758, 62.717, 10.507, 10.884, 5057.38, 2511.347, 142.914]
  MoveL 231 to (2186.49, 124.74, 347.83) mm, rotated rx 179.66 ry -40.68 rz -179.78 deg; joints [106.573, 55.069, -145.55, 72.371, 10.824, 1.075, 5064.994, 2426.388, 142.914]
  MoveL 232 to (2188.58, 61.17, 347.57) mm, rotated rx 179.89 ry -39.72 rz -179.93 deg; joints [106.574, 55.358, -145.55, 72.829, 9.779, 0.605, 5059.421, 2368.078, 142.914]
  MoveL 233 to (2189.63, -0.05, 347.57) mm, rotated rx 177.08 ry -39.67 rz -178.14 deg; joints [106.485, 55.315, -145.496, 85.382, 9.976, -12.043, 5059.422, 2287.176, 142.914]
  MoveL 234 to (2188.58, -61.27, 347.57) mm, rotated rx 177.19 ry -39.63 rz -178.21 deg; joints [106.485, 55.386, -145.496, 85.375, 9.913, -12.034, 5058.265, 2227.592, 143.318]
  MoveL 235 to (2186.49, -124.84, 347.83) mm, rotated rx 178.12 ry -40.61 rz -178.77 deg; joints [106.485, 56.321, -145.496, 85.442, 10.624, -12.137, 5068.383, 2182.492, 152.422]
  MoveL 236 to (2183.35, -193.12, 348.09) mm, rotated rx 174.61 ry -39.89 rz -176.54 deg; joints [106.485, 56.4, -145.496, 100.358, 10.957, -27.291, 5060.002, 2090.503, 152.422]
  MoveL 237 to (2178.9, -262.97, 348.88) mm, rotated rx 174.3 ry -39.37 rz -176.38 deg; joints [106.485, 56.637, -145.496, 104.133, 10.693, -31.088, 5051.771, 2021.033, 152.422]
  MoveL 238 to (2173.41, -330.47, 349.66) mm, rotated rx 175.4 ry -39.48 rz -177.07 deg; joints [106.485, 57.487, -145.496, 104.431, 10.519, -31.391, 5049.97, 1971.867, 157.986]
  MoveL 239 to (2166.87, -388.81, 350.45) mm, rotated rx 172.81 ry -40.11 rz -175.35 deg; joints [106.485, 57.194, -145.132, 110.56, 12.258, -37.75, 5050.101, 1894.984, 157.986]
  MoveL 240 to (2160.33, -431.97, 351.49) mm, rotated rx 166.01 ry -40.37 rz -170.84 deg; joints [106.434, 56.28, -143.996, 123.369, 16.537, -51.125, 5050.101, 1802.95, 157.986]
  MoveL 241 to (2153, -464.41, 352.54) mm, rotated rx 160.9 ry -39.85 rz -167.49 deg; joints [106.434, 55.404, -142.91, 130.35, 19.961, -58.585, 5043.984, 1732.601, 157.986]
  MoveL 242 to (2144.89, -491.88, 353.59) mm, rotated rx 156.15 ry -37.28 rz -165.01 deg; joints [106.434, 54.71, -142.051, 139.84, 23.043, -68.241, 5019.714, 1664.422, 157.986]
  MoveL 243 to (2136, -514.12, 354.9) mm, rotated rx 154.92 ry -35.84 rz -164.67 deg; joints [106.434, 54.699, -142.037, 143.78, 23.876, -72.068, 4999.885, 1629.706, 157.986]
  MoveL 244 to (2127.1, -531.65, 355.94) mm, rotated rx 150.67 ry -31.64 rz -163.57 deg; joints [106.434, 53.624, -140.71, 153.832, 27.755, -81.731, 4959.024, 1566.483, 157.986]
  MoveL 245 to (2117.68, -546.56, 356.99) mm, rotated rx 150.34 ry -30.97 rz -163.66 deg; joints [106.434, 53.627, -140.71, 155.277, 28.128, -83.048, 4943.838, 1547.308, 157.817]
  MoveL 246 to (2107.22, -561.47, 358.3) mm, rotated rx 149.93 ry -30.68 rz -163.54 deg; joints [106.434, 53.62, -140.701, 155.795, 28.518, -83.537, 4931.518, 1528.723, 157.817]
  MoveL 247 to (2096.23, -576.65, 359.6) mm, rotated rx 149.62 ry -28.44 rz -164.4 deg; joints [106.447, 53.702, -140.701, 160.752, 29.3, -87.953, 4899.295, 1505.738, 157.816]
  MoveL 248 to (2084.2, -591.82, 361.17) mm, rotated rx 150.5 ry -29.63 rz -164.37 deg; joints [106.447, 54.289, -140.959, 158.703, 28.608, -86.167, 4898.672, 1505.738, 157.816]
  MoveL 249 to (2071.9, -606.99, 363.01) mm, rotated rx 150.19 ry -30.18 rz -163.93 deg; joints [106.447, 54.367, -140.959, 157.388, 28.836, -85.034, 4892.918, 1491.086, 157.897]
  MoveL 250 to (2059.08, -622.17, 364.84) mm, rotated rx 148.4 ry -29.34 rz -163.23 deg; joints [106.47, 53.784, -140.24, 158.542, 30.649, -86.192, 4875.83, 1458.776, 157.916]
  MoveL 251 to (2046.26, -636.82, 366.67) mm, rotated rx 146.93 ry -28.45 rz -162.77 deg; joints [106.514, 53.286, -139.627, 159.762, 32.212, -87.375, 4857.803, 1429.275, 157.916]
  MoveL 252 to (2033.71, -650.68, 368.76) mm, rotated rx 145.01 ry -26.5 rz -162.65 deg; joints [106.71, 52.474, -138.629, 162.591, 34.552, -90.022, 4831.597, 1392.54, 157.916]
  MoveL 253 to (2014.35, -671.09, 371.9) mm, rotated rx 146.43 ry -25.93 rz -163.82 deg; joints [106.71, 53.433, -138.629, 164.887, 34.44, -92.051, 4805.986, 1392.54, 156.412]
  MoveL 254 to (1994.72, -691.23, 375.3) mm, rotated rx 150.12 ry -25.96 rz -165.88 deg; joints [106.719, 55.682, -141.397, 166.739, 30.771, -93.564, 4780.125, 1407.538, 156.409]
  MoveL 255 to (1981.12, -704.84, 377.39) mm, rotated rx 151.4 ry -25.12 rz -166.97 deg; joints [106.79, 56.236, -141.475, 169.359, 30.418, -95.953, 4757.767, 1407.539, 154.325]
  MoveL 256 to (1966.99, -718.44, 379.49) mm, rotated rx 151.39 ry -23.39 rz -167.78 deg; joints [107.001, 56.382, -141.475, 172.749, 31.181, -99.048, 4728.669, 1391.524, 154.325]
  MoveL 257 to (1952.34, -731.78, 381.58) mm, rotated rx 152.53 ry -23.42 rz -168.32 deg; joints [107.001, 57.134, -142.133, 173.489, 30.302, -99.759, 4713.498, 1391.525, 154.325]
  MoveL 258 to (1937.43, -745.13, 383.93) mm, rotated rx 154.59 ry -22.91 rz -169.52 deg; joints [107.001, 58.231, -143.49, 176.038, 28.494, -102.105, 4690.697, 1397.136, 154.325]
  MoveL 259 to (1922.26, -758.21, 386.55) mm, rotated rx 155.45 ry -21.58 rz -170.46 deg; joints [107.146, 58.765, -143.49, 179.396, 28.867, -105.249, 4664.234, 1394.894, 154.325]
  MoveL 260 to (1906.56, -770.76, 389.17) mm, rotated rx 154.41 ry -20.18 rz -170.62 deg; joints [107.434, 58.509, -143.173, 181.082, 30.425, -106.829, 4638.778, 1370.419, 154.325]
  MoveL 261 to (1889.56, -782.54, 392.31) mm, rotated rx 152.43 ry -19.85 rz -169.95 deg; joints [107.616, 57.998, -142.54, 179.949, 32.348, -105.768, 4623.007, 1340.119, 154.342]
  MoveL 262 to (1871.24, -793.79, 395.97) mm, rotated rx 150.88 ry -17.59 rz -170.44 deg; joints [108.21, 57.373, -141.764, 182.312, 34.872, -107.974, 4589.417, 1309.873, 154.342]
  MoveL 263 to (1851.1, -803.73, 400.15) mm, rotated rx 150.1 ry -17.68 rz -170.09 deg; joints [108.25, 57.509, -141.764, 181.501, 35.612, -107.22, 4572.522, 1295.371, 154.341]
  MoveL 264 to (1827.55, -813.67, 405.91) mm, rotated rx 149.79 ry -15.7 rz -171.05 deg; joints [108.816, 57.649, -141.764, 184.163, 37.021, -109.732, 4535.056, 1280.972, 154.341]
  MoveL 265 to (1801.39, -821.26, 419.78) mm, rotated rx 149.82 ry -24.63 rz -166.38 deg; joints [106.405, 60.47, -145.263, 169.842, 32.377, -96.011, 4579.661, 1304.114, 154.34]
  MoveL 266 to (1776.02, -827.01, 435.21) mm, rotated rx 148.97 ry -27.45 rz -164.51 deg; joints [105.816, 61.142, -145.967, 164.194, 32.191, -90.708, 4579.661, 1304.114, 147.248]
  MoveL 267 to (1751.16, -831.46, 451.69) mm, rotated rx 150.1 ry -28.63 rz -164.6 deg; joints [105.816, 62.355, -147.484, 162.159, 30.629, -88.887, 4564.98, 1314.268, 137.157]
  MoveL 268 to (1726.57, -834.86, 468.7) mm, rotated rx 150.49 ry -30.7 rz -163.88 deg; joints [105.816, 63.525, -148.951, 157.704, 29.585, -84.931, 4560.914, 1322.584, 129.752]
  MoveL 269 to (1702.76, -837.74, 485.44) mm, rotated rx 151.86 ry -30.15 rz -164.96 deg; joints [106.009, 64.103, -149.678, 159.192, 28.378, -86.314, 4530.959, 1328.381, 113.089]
  MoveL 270 to (1680.26, -840.35, 499.83) mm, rotated rx 154.09 ry -27.52 rz -167.35 deg; joints [106.771, 64.388, -150.037, 165.571, 26.992, -92.615, 4486.11, 1333.324, 93.065]
  MoveL 271 to (1658.81, -843.75, 509.77) mm, rotated rx 157.01 ry -21.84 rz -171.03 deg; joints [108.173, 64.388, -150.037, 179.324, 26.525, -106.294, 4418.186, 1337.761, 75.545]
  MoveL 272 to (1639.45, -846.89, 516.83) mm, rotated rx 159.1 ry -18.25 rz -173.18 deg; joints [108.936, 64.513, -150.195, 188.37, 26.605, -115.311, 4368.679, 1345.702, 66.85]
  MoveL 273 to (1621.4, -849.51, 523.37) mm, rotated rx 158.95 ry -19.83 rz -172.56 deg; joints [108.936, 64.98, -150.565, 184.925, 25.978, -112.226, 4367.349, 1345.702, 63.218]
  MoveL 274 to (1598.64, -851.86, 533.05) mm, rotated rx 163.1 ry -20.89 rz -173.82 deg; joints [108.936, 67.313, -153.524, 187.614, 21.485, -115.312, 4352.071, 1383.742, 63.218]
  MoveL 275 to (1578.5, -852.13, 544.3) mm, rotated rx 166.36 ry -25.18 rz -174.1 deg; joints [108.104, 69.412, -156.211, 180.65, 16.204, -108.297, 4362.266, 1421.135, 63.218]
  MoveL 276 to (1564.89, -851.08, 552.68) mm, rotated rx 164.48 ry -25.95 rz -173.07 deg; joints [108.104, 69.923, -156.211, 175.998, 17.982, -103.752, 4359.655, 1412.797, 63.218]
  Set speed (1000.0 mm/s)
  MoveL 277 to (1564.89, -851.08, 552.68) mm, rotated rx 164.48 ry -25.95 rz -173.07 deg; joints [108.104, 69.923, -156.211, 175.998, 17.982, -103.752, 4359.655, 1412.797, 63.218]
  MoveL 278 to (1609.98, -872.56, 639.31) mm, rotated rx 164.48 ry -25.95 rz -173.07 deg; joints [108.046, 72.408, -156.773, 176.413, 19.9, -104.129, 4411.021, 1412.797, 0.001]
  Set speed (1000.0 mm/s)
  MoveL 279 to (1864.64, -820.2, 519.36) mm, rotated rx 168.26 ry -50.58 rz -170.88 deg; joints [108.06, 67.965, -156.773, 93.276, 22.414, -22.96, 4872.798, 1487.01, 123.741]
  MoveL 280 to (1786.74, -812.1, 457.19) mm, rotated rx 168.26 ry -50.58 rz -170.88 deg; joints [108.06, 67.965, -156.773, 93.276, 22.414, -22.96, 4794.897, 1495.108, 185.917]
  MoveL 281 to (1786.74, -812.1, 457.19) mm, rotated rx 168.26 ry -50.58 rz -170.88 deg; joints [108.06, 67.965, -156.773, 93.276, 22.414, -22.96, 4794.897, 1495.108, 185.917]
  Set speed (200.0 mm/s)
  MoveL 282 to (1808.46, -807.91, 444.37) mm, rotated rx 168.26 ry -50.58 rz -170.88 deg; joints [108.06, 67.964, -156.773, 93.274, 22.414, -22.958, 4816.608, 1499.283, 198.727]
  MoveL 283 to (1829.65, -801.9, 432.59) mm, rotated rx 170.89 ry -51.35 rz -172.86 deg; joints [108.061, 67.964, -156.773, 88.778, 22.348, -18.163, 4842.365, 1520.223, 211.094]
  MoveL 284 to (1849.53, -794.57, 422.65) mm, rotated rx 172.79 ry -51.65 rz -174.33 deg; joints [108.061, 67.353, -156.773, 84.329, 22.233, -13.366, 4861.458, 1531.218, 215.503]
  MoveL 285 to (1868.1, -785.94, 414.8) mm, rotated rx 174.14 ry -50.42 rz -175.48 deg; joints [108.061, 67.129, -156.773, 82.7, 20.844, -11.502, 4868.26, 1543.27, 215.509]
  MoveL 286 to (1885.11, -775.73, 408.79) mm, rotated rx 175.21 ry -51.64 rz -176.24 deg; joints [108.061, 67.129, -156.773, 80.214, 21.87, -8.913, 4895.186, 1560.187, 226.074]
  MoveL 287 to (1901.07, -764.48, 404.34) mm, rotated rx 177.95 ry -50.11 rz -178.43 deg; joints [108.061, 67.427, -157.158, 76.231, 20.103, -4.571, 4897.605, 1585.732, 226.074]
  MoveL 288 to (1916.24, -752.45, 400.94) mm, rotated rx 165.53 ry -48.63 rz -169.04 deg; joints [107.147, 66.611, -156.107, 99.049, 21.729, -27.932, 4897.605, 1529.438, 226.074]
  MoveL 289 to (1930.63, -740.42, 398.06) mm, rotated rx 164.44 ry -49.01 rz -168.13 deg; joints [107.147, 66.123, -156.107, 98.6, 22.39, -27.547, 4914.819, 1531.209, 227.769]
  MoveL 290 to (1944.49, -728.38, 395.45) mm, rotated rx 162.57 ry -49.09 rz -166.66 deg; joints [107.059, 65.48, -155.486, 100.715, 23.219, -29.816, 4929.865, 1531.209, 227.769]
  MoveL 291 to (1957.58, -716.09, 393.35) mm, rotated rx 158.8 ry -50.02 rz -163.44 deg; joints [107.013, 64.241, -153.902, 103.601, 25.668, -33.311, 4954.972, 1524.879, 228.71]
  MoveL 292 to (1969.61, -703.27, 392.31) mm, rotated rx 155.21 ry -47.77 rz -161.12 deg; joints [107.013, 64.089, -153.707, 110.699, 26.151, -40.775, 4954.442, 1511.813, 228.71]
  MoveL 293 to (1980.07, -689.4, 393.09) mm, rotated rx 153.94 ry -42.95 rz -161.57 deg; joints [107.013, 65.074, -153.707, 123.721, 25.213, -53.65, 4929.308, 1511.813, 226.345]
  MoveL 294 to (1988.97, -674.23, 395.97) mm, rotated rx 151.38 ry -39.8 rz -160.74 deg; joints [107.013, 65.287, -153.707, 132.317, 26.337, -62.191, 4916.601, 1502.884, 226.345]
  MoveL 295 to (1996.29, -658.01, 400.42) mm, rotated rx 149.14 ry -38.48 rz -159.6 deg; joints [106.926, 65.202, -153.599, 135.776, 27.863, -65.672, 4916.601, 1501.19, 226.345]
  MoveL 296 to (2002.83, -641.26, 405.91) mm, rotated rx 147.45 ry -36.38 rz -159.26 deg; joints [106.929, 65.348, -153.599, 140.694, 29.171, -70.458, 4908.74, 1501.19, 225.442]
  MoveL 297 to (2007.81, -626.88, 410.88) mm, rotated rx 145.73 ry -33 rz -159.64 deg; joints [106.99, 65.477, -153.599, 147.892, 30.816, -77.206, 4887.443, 1493.079, 225.441]
  MoveL 298 to (2008.85, -624.78, 411.4) mm, rotated rx 145.8 ry -32.43 rz -159.98 deg; joints [107.129, 65.493, -153.599, 149.029, 30.836, -78.329, 4884.268, 1493.078, 224.508]
  MoveL 299 to (2010.16, -622.69, 411.67) mm, rotated rx 144.92 ry -31.6 rz -159.8 deg; joints [107.195, 65.164, -153.18, 150.534, 31.757, -79.82, 4880.525, 1485.708, 224.508]
  MoveL 300 to (2011.73, -620.86, 411.4) mm, rotated rx 144.59 ry -30.88 rz -159.96 deg; joints [107.337, 65.003, -152.975, 151.825, 32.186, -81.107, 4877.392, 1481.956, 224.508]
  MoveL 301 to (2024.55, -604.9, 409.83) mm, rotated rx 145.21 ry -30.45 rz -160.61 deg; joints [107.337, 65.083, -153.077, 152.975, 31.718, -82.041, 4883.984, 1500.34, 224.093]
  MoveL 302 to (2039.72, -586.06, 408) mm, rotated rx 143.8 ry -30.75 rz -159.48 deg; joints [107.117, 64.154, -153.077, 151.266, 32.046, -80.28, 4901.128, 1501.888, 224.095]
  MoveL 303 to (2053.33, -568.27, 406.69) mm, rotated rx 143.35 ry -30.75 rz -159.17 deg; joints [107.099, 63.766, -153.077, 150.815, 32.088, -79.823, 4914.619, 1512.61, 224.095]
  MoveL 304 to (2064.84, -551.53, 406.17) mm, rotated rx 140.26 ry -29.2 rz -157.92 deg; joints [107.099, 62.136, -151.01, 152.957, 35.386, -82.054, 4919.825, 1500.879, 224.096]
  MoveL 305 to (2073.47, -536.1, 406.96) mm, rotated rx 141.5 ry -28.05 rz -159.49 deg; joints [107.758, 62.24, -151.141, 155.232, 34.555, -84.404, 4918.999, 1517.394, 218.647]
  MoveL 306 to (2079.75, -522.23, 408.79) mm, rotated rx 142.14 ry -29.17 rz -159.25 deg; joints [107.425, 62.799, -151.849, 153.479, 33.631, -82.562, 4931.702, 1541.857, 218.647]
  MoveL 307 to (2083.94, -508.89, 411.14) mm, rotated rx 142.39 ry -28.01 rz -160.11 deg; joints [108.409, 62.371, -151.844, 154.756, 33.282, -84.369, 4931.698, 1544.297, 211.833]
  MoveL 308 to (2086.55, -494.5, 414.8) mm, rotated rx 144.01 ry -27.32 rz -161.57 deg; joints [108.847, 62.927, -152.549, 156.52, 31.914, -86.13, 4926.814, 1566.478, 206.049]
  MoveL 309 to (2088.12, -477.23, 420.04) mm, rotated rx 145.02 ry -26.19 rz -162.84 deg; joints [109.403, 62.959, -152.59, 158.925, 31.322, -88.635, 4919.325, 1584.99, 197.053]
  MoveL 310 to (2088.38, -459.44, 425.79) mm, rotated rx 145.62 ry -26.52 rz -163.01 deg; joints [109.298, 63.458, -153.224, 158.547, 30.587, -88.183, 4920.696, 1609.417, 193.074]
  MoveL 311 to (2087.6, -443.22, 431.55) mm, rotated rx 146.95 ry -26.53 rz -163.79 deg; joints [109.375, 64.216, -154.191, 159.037, 29.242, -88.619, 4917.733, 1636.184, 188.621]
  MoveL 312 to (2086.29, -429.62, 436.52) mm, rotated rx 144.12 ry -26.95 rz -161.85 deg; joints [108.836, 63.435, -153.195, 157.28, 31.784, -86.738, 4922.72, 1632.123, 188.621]
  MoveL 313 to (2084.72, -419.68, 440.44) mm, rotated rx 143.66 ry -26.54 rz -161.8 deg; joints [109.113, 63.03, -153.195, 157.386, 31.91, -86.998, 4919.554, 1632.189, 183.599]
  MoveL 314 to (2083.15, -411.31, 443.84) mm, rotated rx 141.76 ry -26.34 rz -160.73 deg; joints [108.931, 62.421, -152.42, 157.063, 33.756, -86.668, 4919.554, 1626.789, 183.598]
  MoveL 315 to (2088.12, -379.13, 443.32) mm, rotated rx 140.16 ry -26.15 rz -159.81 deg; joints [108.872, 61.184, -152.42, 155.897, 34.055, -85.436, 4922.554, 1634.288, 182.017]
  MoveL 316 to (2095.18, -319.22, 442.27) mm, rotated rx 139.47 ry -25.88 rz -159.54 deg; joints [108.873, 60.516, -152.42, 155.68, 34.113, -85.133, 4926.495, 1681.234, 181.423]
  MoveL 317 to (2100.42, -260.09, 441.49) mm, rotated rx 139.47 ry -25.87 rz -159.54 deg; joints [108.873, 60.413, -152.421, 155.641, 34.024, -85.077, 4931.193, 1739.092, 181.424]
  MoveL 318 to (2105.13, -193.12, 440.7) mm, rotated rx 137.61 ry -24.56 rz -159.22 deg; joints [109.361, 58.284, -152.42, 155.529, 34.055, -84.959, 4924.516, 1763.469, 176.837]
  MoveL 319 to (2108.79, -132.69, 440.18) mm, rotated rx 137.02 ry -24.42 rz -158.93 deg; joints [109.361, 57.764, -152.42, 155.155, 34.135, -84.545, 4926.743, 1813.686, 176.838]
  MoveL 320 to (2110.62, -92.92, 439.92) mm, rotated rx 139.49 ry -25.11 rz -160.07 deg; joints [109.306, 59.242, -154.306, 154.856, 31.418, -84.085, 4927.929, 1875.514, 176.831]
  MoveL 321 to (2111.4, -63.36, 439.66) mm, rotated rx 149.73 ry -27.95 rz -164.7 deg; joints [109.305, 64.262, -160.792, 150.565, 20.608, -79.649, 4932.316, 1994.368, 176.831]
  MoveL 322 to (2111.4, -63.36, 439.66) mm, rotated rx 142.7 ry -44.91 rz -151.73 deg; joints [106.717, 60.75, -160.792, 105.259, 28.788, -34.351, 5074.364, 1994.368, 196.285]
  MoveL 323 to (2119.78, -59.7, 429.72) mm, rotated rx 141.26 ry -45.36 rz -150.28 deg; joints [106.491, 60.443, -160.417, 105.537, 29.93, -34.688, 5088.651, 1994.368, 209.694]
  MoveL 324 to (2127.89, -55.77, 419.51) mm, rotated rx 140.78 ry -45.79 rz -149.67 deg; joints [106.491, 60.245, -160.417, 104.653, 30.414, -33.858, 5101.092, 1996.587, 221.238]
  MoveL 325 to (2136.78, -51.85, 408.79) mm, rotated rx 140.98 ry -46.05 rz -149.74 deg; joints [106.491, 60.246, -160.42, 104.068, 30.432, -33.252, 5111.464, 2002.763, 231.759]
  MoveL 326 to (2140.18, -49.76, 404.6) mm, rotated rx 141.16 ry -49.37 rz -148.57 deg; joints [106.491, 60.246, -160.42, 98.355, 32.252, -27.616, 5140.05, 2024.406, 242.866]
  MoveL 327 to (2142.54, -46.88, 401.72) mm, rotated rx 142.58 ry -50.84 rz -149.32 deg; joints [106.49, 60.246, -160.42, 95.334, 32.425, -24.371, 5149.334, 2040.364, 244.817]
  MoveL 328 to (2142.54, -46.88, 401.72) mm, rotated rx -180 ry -44.31 rz 180 deg; joints [109.67, 69.214, -172.464, 37.522, 22.465, 34.389, 5074.435, 2222.368, 244.817]
  MoveL 329 to (2144.11, -43.48, 399.89) mm, rotated rx 180 ry -44.31 rz -180 deg; joints [109.67, 69.214, -172.464, 37.522, 22.465, 34.389, 5076.005, 2225.768, 246.649]
  MoveL 330 to (2144.63, -39.81, 399.11) mm, rotated rx -180 ry -44.31 rz -180 deg; joints [109.67, 69.214, -172.465, 37.521, 22.466, 34.39, 5076.527, 2229.426, 247.432]
  MoveL 331 to (2144.37, -24.12, 399.11) mm, rotated rx 180 ry -45.71 rz -180 deg; joints [109.67, 69.139, -172.465, 39.383, 23.69, 32.695, 5088.41, 2244.375, 251.5]
  MoveL 332 to (2144.37, -12.08, 399.11) mm, rotated rx 178.57 ry -46.1 rz -178.97 deg; joints [109.543, 68.771, -172.465, 41.456, 23.793, 30.744, 5089.513, 2244.375, 250.396]
  MoveL 333 to (2144.37, -0.05, 399.11) mm, rotated rx 175.75 ry -49.13 rz -176.78 deg; joints [109.439, 68.3, -171.812, 48.808, 25.628, 23.565, 5115.412, 2241.121, 257.486]
  MoveL 334 to (2144.37, 11.99, 399.11) mm, rotated rx -179.73 ry -49.56 rz 179.8 deg; joints [109.439, 68.299, -171.815, 43.542, 27.187, 29.265, 5118.426, 2278.553, 258.299]
  MoveL 335 to (2144.37, 24.28, 399.11) mm, rotated rx 179.8 ry -50.65 rz -179.84 deg; joints [109.439, 68.299, -171.815, 45.207, 28.014, 27.685, 5127.783, 2288.262, 262.74]
  MoveL 336 to (2144.63, 39.98, 399.11) mm, rotated rx -177.81 ry -51.25 rz 178.29 deg; joints [109.439, 68.299, -171.815, 43.263, 29.232, 29.929, 5133.294, 2316.679, 265.467]
  MoveL 337 to (2144.11, 43.64, 399.89) mm, rotated rx -177.4 ry -50.59 rz 177.99 deg; joints [109.439, 68.333, -171.863, 42.103, 28.805, 31.046, 5127.198, 2322.78, 262.346]
  MoveL 338 to (2142.54, 47.04, 401.72) mm, rotated rx -176.05 ry -51.85 rz 176.89 deg; joints [109.439, 68.333, -171.863, 42.192, 30.302, 31.255, 5136.672, 2332.673, 266.269]
  MoveL 339 to (2140.18, 49.66, 404.6) mm, rotated rx -177.95 ry -50.11 rz 178.43 deg; joints [109.439, 68.333, -171.863, 42.141, 28.226, 30.896, 5119.121, 2325.996, 255.568]
  MoveL 340 to (2136.78, 52.01, 408.79) mm, rotated rx 180 ry -45.71 rz -180 deg; joints [109.439, 68.336, -171.863, 39.222, 23.812, 33.116, 5077.288, 2317.144, 234.789]
  MoveL 341 to (2127.89, 55.94, 419.51) mm, rotated rx -178.57 ry -46.11 rz 178.97 deg; joints [109.443, 69.11, -172.938, 37.459, 24.928, 35.068, 5072.33, 2330.474, 233.538]
  MoveL 342 to (2119.78, 59.6, 429.72) mm, rotated rx -175.76 ry -49.16 rz 176.79 deg; joints [109.443, 69.11, -172.938, 38.334, 28.448, 34.826, 5091.328, 2349.24, 235.325]
  MoveL 343 to (2111.4, 63.26, 439.66) mm, rotated rx 179.73 ry -49.56 rz -179.8 deg; joints [109.443, 69.11, -172.937, 43.745, 27.252, 29.062, 5085.74, 2327.567, 226.087]
  MoveL 344 to (2111.4, 63.26, 439.66) mm, rotated rx -134.57 ry -75.84 rz 135.45 deg; joints [109.443, 69.112, -172.939, 53.777, 58.066, 27.444, 5303.441, 2382.918, 413.823]
  MoveL 345 to (2110.62, 92.82, 439.92) mm, rotated rx -124.48 ry -74.06 rz 125.53 deg; joints [109.443, 69.112, -172.94, 52.275, 59.756, 30.569, 5307.218, 2427.082, 423.368]
  MoveL 346 to (2108.79, 132.85, 440.18) mm, rotated rx -114.02 ry -68.32 rz 115.63 deg; joints [109.443, 69.112, -172.94, 48.303, 62.1, 37.642, 5305.352, 2500.682, 432.931]
  MoveL 347 to (2105.13, 193.28, 440.7) mm, rotated rx -111.26 ry -65.32 rz 113.19 deg; joints [109.443, 69.112, -172.94, 46.352, 63.17, 41.002, 5300.257, 2577.603, 436.562]
  MoveL 348 to (2100.42, 260, 441.49) mm, rotated rx -106 ry -60.62 rz 108.21 deg; joints [109.55, 70.876, -175.415, 43.873, 66.44, 46.515, 5300.257, 2667.706, 470.632]
  MoveL 349 to (2095.18, 319.38, 442.27) mm, rotated rx -104.15 ry -54.09 rz 107.29 deg; joints [109.55, 70.876, -175.415, 39.976, 68.817, 53.039, 5288.551, 2761.612, 479.747]
  MoveL 350 to (2088.12, 379.29, 443.32) mm, rotated rx -104.19 ry -49.35 rz 108.44 deg; joints [109.55, 70.876, -175.415, 36.556, 70.197, 57.644, 5271.266, 2849.964, 482.272]
  MoveL 351 to (2083.15, 411.21, 443.84) mm, rotated rx 116.95 ry -61.96 rz -119.95 deg; joints [109.55, 70.876, -175.415, 80.647, 52.175, -13.976, 5256.62, 2536.889, 427.368]
  MoveL 352 to (2084.72, 419.58, 440.44) mm, rotated rx 117.68 ry -64.42 rz -120.18 deg; joints [109.55, 70.876, -175.415, 78.438, 52.847, -10.954, 5264.192, 2560.552, 432.536]
  MoveL 353 to (2086.29, 429.52, 436.52) mm, rotated rx 122.82 ry -71.24 rz -124.26 deg; joints [109.55, 70.876, -175.415, 72.58, 54.415, -2.381, 5277.53, 2611.627, 439.224]
  MoveL 354 to (2087.6, 443.12, 431.55) mm, rotated rx 137.63 ry -75.76 rz -138.52 deg; joints [109.549, 71.231, -175.918, 67.574, 54.381, 5.314, 5277.855, 2657.715, 439.224]
  MoveL 355 to (2088.38, 459.34, 425.79) mm, rotated rx -134.42 ry -73 rz 135.7 deg; joints [109.55, 71.473, -176.262, 50.659, 57.548, 31.202, 5270.52, 2793.795, 439.185]
  MoveL 356 to (2088.12, 477.13, 420.04) mm, rotated rx -116.56 ry -58.51 rz 120.38 deg; joints [109.55, 71.494, -176.273, 38.614, 62.099, 48.733, 5251.278, 2906.825, 454.348]
  MoveL 357 to (2086.55, 494.4, 414.8) mm, rotated rx -109.9 ry -44.97 rz 117.12 deg; joints [109.55, 71.494, -176.273, 29.136, 68.487, 62.174, 5227.639, 3009.628, 489.119]
  MoveL 358 to (2083.94, 508.79, 411.14) mm, rotated rx -105.78 ry -32.39 rz 117.81 deg; joints [109.55, 71.494, -176.273, 20.944, 75.897, 72.672, 5195.292, 3102.605, 537.063]
  MoveL 359 to (2079.75, 522.13, 408.79) mm, rotated rx -104.76 ry -26.01 rz 121 deg; joints [109.55, 70.747, -176.273, 15.285, 80.25, 77.478, 5156.824, 3154.501, 556.567]
  MoveL 360 to (2073.47, 536.26, 406.96) mm, rotated rx -104.78 ry -21.87 rz 125.3 deg; joints [107.732, 68.785, -176.273, 11.519, 84.079, 80.912, 5090.604, 3190.652, 556.568]
  MoveL 361 to (2064.84, 551.43, 406.17) mm, rotated rx -105.02 ry -19.59 rz 128.67 deg; joints [105.422, 67.917, -176.273, 9.819, 85.791, 82.845, 5030.014, 3224.834, 556.571]
  MoveL 362 to (2053.33, 568.18, 406.69) mm, rotated rx -105.8 ry -19.22 rz 130.68 deg; joints [103.673, 67.54, -176.273, 9.53, 85.675, 83.529, 4986.383, 3248.84, 548.713]
  MoveL 363 to (2039.72, 586.23, 408) mm, rotated rx -105.46 ry -17.68 rz 132.32 deg; joints [102.793, 66.56, -176.273, 8.291, 87.671, 84.579, 4946.598, 3270.544, 548.713]
  MoveL 364 to (2024.55, 604.8, 409.83) mm, rotated rx -104.64 ry -16.7 rz 132.26 deg; joints [102.957, 66.56, -176.273, 7.842, 88.83, 84.96, 4931.188, 3293.634, 556.449]
  MoveL 365 to (2011.73, 620.76, 411.4) mm, rotated rx -105.04 ry -17.29 rz 132.12 deg; joints [103.317, 65.945, -176.273, 7.842, 88.829, 84.676, 4922.273, 3299.113, 546.109]
  MoveL 366 to (2010.16, 622.85, 411.67) mm, rotated rx -104.76 ry -21.4 rz 125.83 deg; joints [107.86, 67.646, -176.273, 10.737, 85.458, 81.332, 5019.976, 3269.529, 546.109]
  MoveL 367 to (2008.85, 624.95, 411.4) mm, rotated rx -105.15 ry -23.35 rz 124.34 deg; joints [108.128, 68.942, -176.266, 12.589, 82.926, 79.934, 5039.656, 3269.069, 546.116]
  MoveL 368 to (2007.81, 627.04, 410.88) mm, rotated rx -107.65 ry -27.86 rz 124.25 deg; joints [108.127, 68.942, -176.266, 14.805, 78.934, 77.126, 5049.117, 3245.393, 516.718]
  MoveL 369 to (2002.83, 641.17, 405.91) mm, rotated rx -107.93 ry -28.38 rz 124.25 deg; joints [108.415, 68.503, -176.266, 14.805, 78.934, 76.811, 5046.463, 3251.147, 515.633]
  MoveL 370 to (1996.29, 657.91, 400.42) mm, rotated rx -109.04 ry -27.49 rz 126.78 deg; joints [106.424, 68.256, -176.266, 14.147, 78.627, 78.024, 5003.264, 3282.204, 513.531]
  MoveL 371 to (1988.97, 674.13, 395.97) mm, rotated rx -109.01 ry -24.18 rz 130.06 deg; joints [104.944, 66.24, -176.266, 11.098, 82.092, 80.815, 4946.32, 3308.515, 513.531]
  MoveL 372 to (1980.07, 689.3, 393.09) mm, rotated rx -108.69 ry -20.6 rz 133.88 deg; joints [102.797, 63.714, -176.266, 8.134, 86.473, 83.558, 4875.442, 3329.885, 513.532]
  MoveL 373 to (1969.61, 703.17, 392.31) mm, rotated rx -110.28 ry -18.9 rz 138.76 deg; joints [98.303, 63.395, -176.266, 7.27, 86.188, 85.667, 4785.71, 3362.997, 505.162]
  MoveL 374 to (1957.58, 715.99, 393.35) mm, rotated rx -108.98 ry -16.34 rz 140.71 deg; joints [97.473, 60.594, -176.266, 5.244, 91.292, 86.972, 4739.576, 3363.02, 507.061]
  MoveL 375 to (1944.49, 728.28, 395.45) mm, rotated rx -107.25 ry -14.65 rz 140.84 deg; joints [97.473, 60.594, -176.266, 4.484, 93.573, 87.42, 4720.636, 3385.544, 523.844]
  MoveL 376 to (1930.63, 740.32, 398.06) mm, rotated rx -106.75 ry -13.85 rz 141.5 deg; joints [96.9, 60.545, -176.266, 4.139, 94.423, 87.777, 4694.778, 3402.612, 527.497]
  MoveL 377 to (1916.24, 752.61, 400.94) mm, rotated rx -104.52 ry -11.48 rz 142.45 deg; joints [96.242, 60.491, -176.266, 3.116, 97.54, 88.436, 4661.373, 3428.373, 550.37]
  MoveL 378 to (1901.07, 764.39, 404.34) mm, rotated rx -104.71 ry -10.88 rz 144.27 deg; joints [94.387, 60.596, -176.416, 2.995, 97.704, 89.029, 4615.082, 3446.162, 548.563]
  MoveL 379 to (1885.11, 775.64, 408.79) mm, rotated rx -105.46 ry -10.29 rz 147.13 deg; joints [91.558, 60.276, -176.416, 2.815, 97.662, 89.881, 4551.177, 3459.003, 538.521]
  MoveL 380 to (1868.1, 785.84, 414.8) mm, rotated rx -105.4 ry -8.87 rz 150.78 deg; joints [87.927, 60.328, -176.495, 2.425, 98.425, 90.987, 4471.127, 3476.042, 538.521]
  MoveL 381 to (1849.53, 794.47, 422.65) mm, rotated rx -105.79 ry -7.76 rz 154.48 deg; joints [84.141, 60.502, -176.743, 2.208, 98.704, 92.099, 4388.261, 3485.885, 533.269]
  MoveL 382 to (1829.65, 802.06, 432.59) mm, rotated rx -107.79 ry -8.17 rz 156.11 deg; joints [82.345, 60.473, -176.743, 2.41, 96.791, 92.839, 4341.715, 3485.886, 505.361]
  MoveL 383 to (1808.46, 807.81, 444.37) mm, rotated rx -112.15 ry -9.63 rz 157.65 deg; joints [80.557, 60.473, -176.743, 2.871, 92.311, 93.955, 4298.504, 3473.764, 453.819]
  MoveL 384 to (1786.74, 812.26, 457.19) mm, rotated rx -118.21 ry -11.24 rz 160.03 deg; joints [78.165, 60.473, -176.743, 3.063, 86.291, 95.732, 4245.735, 3448.171, 389.393]
  MoveL 385 to (1762.67, 814.88, 473.41) mm, rotated rx -119.66 ry -12.67 rz 158.94 deg; joints [79.329, 60.473, -176.743, 3.5, 84.357, 95.302, 4245.451, 3443.792, 358.217]
  MoveL 386 to (1738.34, 816.97, 489.89) mm, rotated rx -125.73 ry -17.3 rz 157.55 deg; joints [80.768, 63.767, -176.743, 5.442, 73.685, 94.31, 4260.275, 3443.792, 304.167]
  MoveL 387 to (1713.23, 819.59, 507.42) mm, rotated rx -134.31 ry -18.96 rz 161.59 deg; joints [78.205, 63.767, -176.743, 4.596, 65.608, 96.777, 4197.017, 3389.939, 229.635]
  MoveL 388 to (1688.11, 818.28, 525.47) mm, rotated rx -132.85 ry -17.47 rz 162.07 deg; joints [77.348, 64.389, -177.634, 4.007, 67.784, 97.509, 4152.087, 3400.473, 229.635]
  Set speed (1000.0 mm/s)
  MoveL 389 to (1688.11, 818.28, 525.47) mm, rotated rx -132.85 ry -17.47 rz 162.07 deg; joints [77.348, 64.389, -177.634, 4.007, 67.784, 97.509, 4152.087, 3400.473, 229.635]
  MoveL 390 to (1730.11, 881.75, 590.34) mm, rotated rx -132.85 ry -17.47 rz 162.07 deg; joints [77.348, 64.389, -177.634, 4.007, 67.784, 97.509, 4194.085, 3463.94, 164.766]

